FUNCTION_BLOCK pump_slider (* Composite Function Block Type *)
  (* Standard: 61499-2 *)
  (* Version 0.0, 12/30/2019, prana, nxtControl GmbH, template *)
  PACKAGE Main;
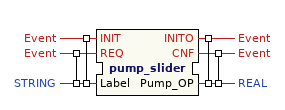
  EVENT_INPUT
    INIT WITH Label; (* Initialization Request *)
    REQ WITH Label; (* Normal Execution Request *)
  END_EVENT
  EVENT_OUTPUT
    INITO WITH Pump_OP; (* Initialization Confirm *)
    CNF WITH Pump_OP; (* Execution Confirmation *)
  END_EVENT
  VAR_INPUT
    Label : STRING; (* Input event qualifier *)
  END_VAR
  VAR_OUTPUT
    Pump_OP : REAL; (* Output event qualifier *)
  END_VAR
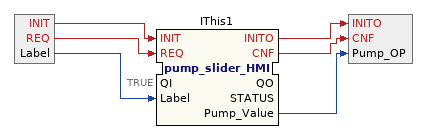
  FBS
    IThis1 : pump_slider_HMI(QI := TRUE);
  END_FBS
  EVENT_CONNECTIONS
    INIT TO IThis1.INIT;
    REQ TO IThis1.REQ;
    IThis1.INITO TO INITO;
    IThis1.CNF TO CNF;
  END_CONNECTIONS
  DATA_CONNECTIONS
    Label TO IThis1.Label;
    IThis1.Pump_Value TO Pump_OP;
  END_CONNECTIONS
END_FUNCTION_BLOCK
